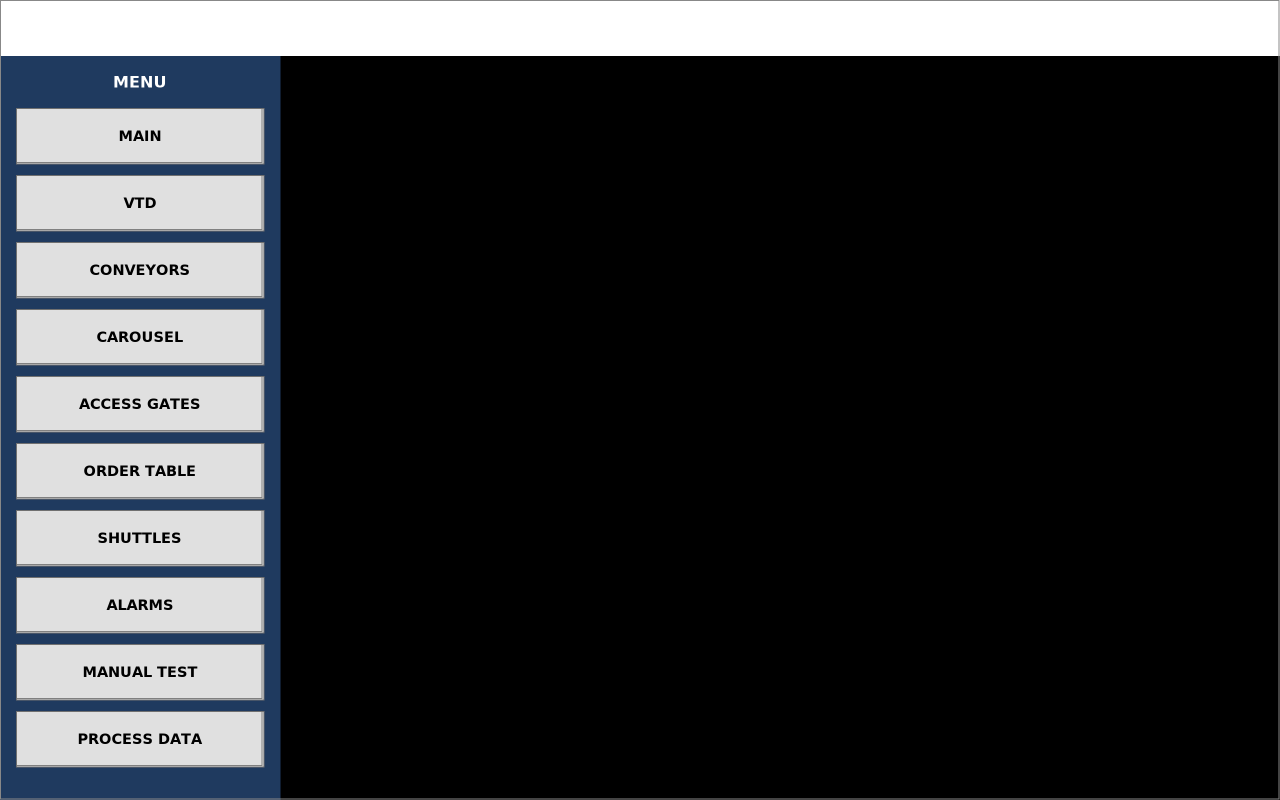
VISUALIZATION Dialog  // 1280x800
    Rectangle (0,0 1280x56)
        OnMouseClick: CloseDialog Dialog=Current Dialog, Result=OK, NumpadKeypadSet=True
    Rectangle (280,56 1000x744)
        OnMouseClick: CloseDialog Dialog=Current Dialog, Result=OK, NumpadKeypadSet=True
    Rectangle (0,56 280x744)
    Rectangle (12,64 256x36), "MENU"
    Button (16,108 248x56), "MAIN"
        OnMouseDown: change screen: Main
        OnMouseClick: CloseDialog Dialog=Current Dialog, Result=OK, NumpadKeypadSet=True
    Button (16,175 248x56), "VTD"
        OnMouseDown: change screen: VTD
        OnMouseClick: CloseDialog Dialog=Current Dialog, Result=OK, NumpadKeypadSet=True
    Button (16,242 248x56), "CONVEYORS"
        OnMouseDown: change screen: CNV
        OnMouseClick: CloseDialog Dialog=Current Dialog, Result=OK, NumpadKeypadSet=True
    Button (16,309 248x56), "CAROUSEL"
        OnMouseDown: change screen: Carrousel
        OnMouseClick: CloseDialog Dialog=Current Dialog, Result=OK, NumpadKeypadSet=True
    Button (16,376 248x56), "ACCESS GATES"
        OnMouseDown: change screen: Access_Gates
        OnMouseClick: CloseDialog Dialog=Current Dialog, Result=OK, NumpadKeypadSet=True
    Button (16,443 248x56), "ORDER TABLE"
        OnMouseDown: change screen: Order_Table
        OnMouseClick: CloseDialog Dialog=Current Dialog, Result=OK, NumpadKeypadSet=True
    Button (16,510 248x56), "SHUTTLES"
        OnMouseDown: change screen: Shuttles
        OnMouseClick: CloseDialog Dialog=Current Dialog, Result=OK, NumpadKeypadSet=True
    Button (16,577 248x56), "ALARMS"
        OnMouseDown: change screen: Alarms
        OnMouseClick: CloseDialog Dialog=Current Dialog, Result=OK, NumpadKeypadSet=True
    Button (16,644 248x56), "MANUAL TEST"
        OnMouseDown: change screen: VTDManualTest
        OnMouseClick: CloseDialog Dialog=Current Dialog, Result=OK, NumpadKeypadSet=True
    Button (16,711 248x56), "PROCESS DATA"
        OnMouseDown: change screen: Visualization
        OnMouseClick: CloseDialog Dialog=Current Dialog, Result=OK, NumpadKeypadSet=True
END_VISUALIZATION

(* stored: Version 1.1.0.1
   Visu Dialog: Id {8067e270-ca00-4168-8692-f5659e66b526} *)
